FUNCTION_BLOCK fbShutterCmdSourceSwitch IMPLEMENTS iShutterCmdSource
VAR_INPUT
    OpenSwitchState : stSwitchState;
    CloseSwitchState : stSwitchState;
    ShutterStateType : eShutterStateType;
END_VAR
VAR PERSISTENT
    OpenLongClickPosition : stShutterPosition := (Height := 50, Angle := 100);
    CloseLongClickPosition : stShutterPosition := (Height := 0, Angle := 100);
END_VAR

METHOD Process
VAR_IN_OUT
	CmdEvent	: stShutterCmdEvent;
END_VAR
VAR
	NewCmd : stShutterCmd;
END_VAR

// Exit if both switches are idle
IF OpenSwitchState.StateType = eSwitchStateType.IDLE AND
   CloseSwitchState.StateType = eSwitchStateType.IDLE THEN
    RETURN;
END_IF

// If shutter is moving and any switch was pressed
IF ShutterStateType <> eShutterStateType.IDLE THEN
    NewCmd.CommandType := eShutterCmdType.STOP;
    CmdEvent.Execute := TRUE;
// Double Open click
ELSIF (OpenSwitchState.StateType = eSwitchStateType.MULTI_CLICK) AND (OpenSwitchState.PressCount = 2) THEN
    NewCmd.CommandType := eShutterCmdType.OPEN;
    CmdEvent.Execute := TRUE;
// Double Close click
ELSIF (CloseSwitchState.StateType = eSwitchStateType.MULTI_CLICK) AND (CloseSwitchState.PressCount = 2) THEN
    NewCmd.CommandType := eShutterCmdType.CLOSE;
    CmdEvent.Execute := TRUE;
// Short Open click
ELSIF OpenSwitchState.StateType = eSwitchStateType.SHORT_CLICK THEN
    NewCmd.CommandType := eShutterCmdType.STEP_OPEN;
    CmdEvent.Execute := TRUE;
// Short Close click
ELSIF CloseSwitchState.StateType = eSwitchStateType.SHORT_CLICK THEN
    NewCmd.CommandType := eShutterCmdType.STEP_CLOSE;
    CmdEvent.Execute := TRUE;
// Long Open click
ELSIF OpenSwitchState.StateType = eSwitchStateType.LONG_CLICK THEN
    NewCmd.CommandType := eShutterCmdType.MOVE_TO_POSITION;
    NewCmd.Position := OpenLongClickPosition;
    CmdEvent.Execute := TRUE;
// Long Close click
ELSIF CloseSwitchState.StateType = eSwitchStateType.LONG_CLICK THEN
    NewCmd.CommandType := eShutterCmdType.MOVE_TO_POSITION;
    NewCmd.Position := CloseLongClickPosition;
    CmdEvent.Execute := TRUE;
END_IF
END_METHOD

END_FUNCTION_BLOCK

(* stored: Version 1.1.0.1
   POU fbShutterCmdSourceSwitch: Id {c862dcf9-c651-483d-a78a-0c62d3a73fd7}, SpecialFunc None
   Method Process: Id {bb7c2f45-924d-4762-a2d7-89765f3d0a73} *)
